// TIA Portal V15.1 export
// export: Created 2026-09-17T17:40:11.6428239Z, ExportSetting WithDefaults, DisplayName Totally Integrated Automation Portal, DisplayVersion V15.1, DisplayName TIA Portal Openness, DisplayVersion V15.1, DisplayName STEP 7 Professional, DisplayVersion V15.1, DisplayName WinCC Professional, DisplayVersion V15.1
Screen "Motion"  1024x768, Number=6
  ScreenLayer 
    Button "Button_1" at 31,675 size 90x44  Mode=Text, StyleItem=Button, TextOff="End RT", TextOn="Text"
      on Press: StopRuntime(Mode := 0)
    GraphicView "Graphic view_1" at 189,10 size 770x758  Picture=images (6)
    Button "Button_2" at 31,619 size 90x44  Mode=Text, StyleItem=Button, TextOff="Back", TextOn="Text"
      on Press: ActivateScreen(Screen name := Start Screen, Object number := 0)
    GraphicView "Graphic view_2" at 818,633 size 158x89  Picture=Graphic_1
    TextField "Text field_1" at 793,722 size 231x21  Text="By Ahmad Saber Zain"
    TextField "Text field_2" at 618,8 size 190x29  Text="Motion Screen"
    GraphicView "Graphic view_9" at 474,348 size 36x30  Picture=Graphic_3
      RangeAppearanceAnimation "RangeAppearanceAnimation"
        tag PLC_1_test1scada
        0..0: back #ffffff, fore #000000
        1..1: back #ffffff, fore #000000, flashing
    GraphicView "Graphic view_3" at 606,193 size 36x30  Picture=Graphic_2
      SingleBitVisibilityAnimation "VisibilityAnimation"  Visible=false
        tag troll_scd_rev_arrow
    GraphicView "Graphic view_4" at 840,191 size 36x30  Picture=Graphic_3
      SingleBitVisibilityAnimation "VisibilityAnimation"  Visible=false
        tag troll_scd_fwd_arrow
    GraphicView "Graphic view_5" at 711,225 size 36x30  Picture=Graphic_4
      SingleBitVisibilityAnimation "VisibilityAnimation"  Visible=false
        tag HYD_scd_up_arrow
    GraphicView "Graphic view_6" at 714,325 size 36x30  Picture=Graphic_5
      SingleBitVisibilityAnimation "VisibilityAnimation"  Visible=false
        tag HYD_scd_down_arrow
    GraphicView "Graphic view_7" at 360,254 size 36x30  Picture=Graphic_2
      SingleBitVisibilityAnimation "VisibilityAnimation"  Visible=false
        tag slewing anticlockwise
    GraphicView "Graphic view_8" at 460,255 size 36x30  Picture=Graphic_3
      RangeAppearanceAnimation "RangeAppearanceAnimation"
        tag slewing clockwise
        0..0: back #ffffff, fore #ffffff
        1..1: back #ffffff, fore #000000, flashing
    TextField "Text field_4" at 264,295 size 167x23  Text="Anti Clockwise"
      SingleBitVisibilityAnimation "VisibilityAnimation"  Visible=false
        tag slewing anticlockwise
    TextField "Text field_5" at 684,355 size 95x23  Text="Down"
      SingleBitVisibilityAnimation "VisibilityAnimation"  Visible=false
        tag HYD_scd_down_arrow
    TextField "Text field_3" at 444,295 size 128x23  Text="Clockwise"
      RangeAppearanceAnimation "RangeAppearanceAnimation"
        tag slewing clockwise
        0..0: back #ffffff, fore #ffffff
        1..1: back #ffffff, fore #000000, flashing
    TextField "Text field_6" at 690,208 size 64x23  Text="UP"
      SingleBitVisibilityAnimation "VisibilityAnimation"  Visible=false
        tag HYD_scd_up_arrow
    TextField "Text field_7" at 825,218 size 97x23  Text="Forward"
      SingleBitVisibilityAnimation "VisibilityAnimation"  Visible=false
        tag troll_scd_fwd_arrow
    TextField "Text field_8" at 578,221 size 111x23  Text="Backward"
      SingleBitVisibilityAnimation "VisibilityAnimation"  Visible=false
        tag troll_scd_rev_arrow
